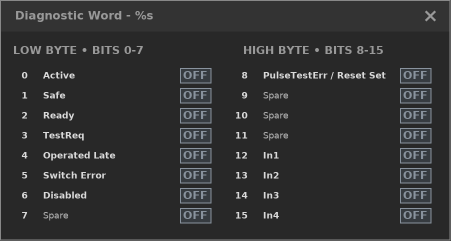
VISUALIZATION FRM_WordDiagnostic  // 451x241
    Rectangle (0,30 451x211)
    Textfield (0,0 411x31), "Diagnostic Word - %s", text variable: Motion_Safety.stSafety.stOut.astDiagnosticElement[GVL_Safety.nHMIDiagWordIndex].sName
    Label (10,40 113x21), "LOW BYTE • BITS 0-7"
    Label (240,40 113x21), "HIGH BYTE • BITS 8-15"
    Label (10,70 21x11), "0"
    Label (10,90 21x11), "1"
    Label (10,110 21x11), "2"
    Label (10,130 21x11), "3"
    Label (10,150 21x11), "4"
    Label (10,170 21x11), "5"
    Label (10,190 21x11), "6"
    Label (10,210 21x11), "7"
    Label (40,70 131x11), "Active"
    Label (40,90 131x11), "Safe"
    Label (40,110 131x11), "Ready"
    Label (40,130 131x11), "TestReq"
    Label (40,150 131x11), "Operated Late"
    Label (40,170 131x11), "Switch Error"
    Label (40,190 131x11), "Disabled"
    Label (40,210 131x11), "Spare"
    Rectangle (180,68 31x15), "ON"
    Rectangle (180,68 31x15), "OFF", invisible if: Motion_Safety.fbMotionSafety.stPNOZEtherCATDiagIn.astDiagnosticElementsIn[GVL_Safety.nHMIDiagWordIndex].nLow.b0
    Rectangle (180,88 31x15), "ON"
    Rectangle (180,88 31x15), "OFF", invisible if: Motion_Safety.fbMotionSafety.stPNOZEtherCATDiagIn.astDiagnosticElementsIn[GVL_Safety.nHMIDiagWordIndex].nLow.b1
    Rectangle (180,108 31x15), "ON"
    Rectangle (180,108 31x15), "OFF", invisible if: Motion_Safety.fbMotionSafety.stPNOZEtherCATDiagIn.astDiagnosticElementsIn[GVL_Safety.nHMIDiagWordIndex].nLow.b2
    Rectangle (180,128 31x15), "ON"
    Rectangle (180,128 31x15), "OFF", invisible if: Motion_Safety.fbMotionSafety.stPNOZEtherCATDiagIn.astDiagnosticElementsIn[GVL_Safety.nHMIDiagWordIndex].nLow.b3
    Rectangle (180,148 31x15), "ON"
    Rectangle (180,148 31x15), "OFF", invisible if: Motion_Safety.fbMotionSafety.stPNOZEtherCATDiagIn.astDiagnosticElementsIn[GVL_Safety.nHMIDiagWordIndex].nLow.b4
    Rectangle (180,168 31x15), "ON"
    Rectangle (180,168 31x15), "OFF", invisible if: Motion_Safety.fbMotionSafety.stPNOZEtherCATDiagIn.astDiagnosticElementsIn[GVL_Safety.nHMIDiagWordIndex].nLow.b5
    Rectangle (180,188 31x15), "ON"
    Rectangle (180,188 31x15), "OFF", invisible if: Motion_Safety.fbMotionSafety.stPNOZEtherCATDiagIn.astDiagnosticElementsIn[GVL_Safety.nHMIDiagWordIndex].nLow.b6
    Rectangle (180,208 31x15), "ON"
    Rectangle (180,208 31x15), "OFF", invisible if: Motion_Safety.fbMotionSafety.stPNOZEtherCATDiagIn.astDiagnosticElementsIn[GVL_Safety.nHMIDiagWordIndex].nLow.b7
    Label (230,70 21x11), "8"
    Label (230,90 21x11), "9"
    Label (230,110 21x11), "10"
    Label (230,130 21x11), "11"
    Label (230,150 21x11), "12"
    Label (230,170 21x11), "13"
    Label (230,190 21x11), "14"
    Label (230,210 21x11), "15"
    Label (260,70 131x11), "PulseTestErr / Reset Set"
    Label (260,90 131x11), "Spare"
    Label (260,110 131x11), "Spare"
    Label (260,130 131x11), "Spare"
    Label (260,150 131x11), "In1"
    Label (260,170 131x11), "In2"
    Label (260,190 131x11), "In3"
    Label (260,210 131x11), "In4"
    Rectangle (400,68 31x15), "ON"
    Rectangle (400,68 31x15), "OFF", invisible if: Motion_Safety.fbMotionSafety.stPNOZEtherCATDiagIn.astDiagnosticElementsIn[GVL_Safety.nHMIDiagWordIndex].nHigh.b0
    Rectangle (400,88 31x15), "ON"
    Rectangle (400,88 31x15), "OFF", invisible if: Motion_Safety.fbMotionSafety.stPNOZEtherCATDiagIn.astDiagnosticElementsIn[GVL_Safety.nHMIDiagWordIndex].nHigh.b1
    Rectangle (400,108 31x15), "ON"
    Rectangle (400,108 31x15), "OFF", invisible if: Motion_Safety.fbMotionSafety.stPNOZEtherCATDiagIn.astDiagnosticElementsIn[GVL_Safety.nHMIDiagWordIndex].nHigh.b2
    Rectangle (400,128 31x15), "ON"
    Rectangle (400,128 31x15), "OFF", invisible if: Motion_Safety.fbMotionSafety.stPNOZEtherCATDiagIn.astDiagnosticElementsIn[GVL_Safety.nHMIDiagWordIndex].nHigh.b3
    Rectangle (400,148 31x15), "ON"
    Rectangle (400,148 31x15), "OFF", invisible if: Motion_Safety.fbMotionSafety.stPNOZEtherCATDiagIn.astDiagnosticElementsIn[GVL_Safety.nHMIDiagWordIndex].nHigh.b4
    Rectangle (400,168 31x15), "ON"
    Rectangle (400,168 31x15), "OFF", invisible if: Motion_Safety.fbMotionSafety.stPNOZEtherCATDiagIn.astDiagnosticElementsIn[GVL_Safety.nHMIDiagWordIndex].nHigh.b5
    Rectangle (400,188 31x15), "ON"
    Rectangle (400,188 31x15), "OFF", invisible if: Motion_Safety.fbMotionSafety.stPNOZEtherCATDiagIn.astDiagnosticElementsIn[GVL_Safety.nHMIDiagWordIndex].nHigh.b6
    Rectangle (400,208 31x15), "ON"
    Rectangle (400,208 31x15), "OFF", invisible if: Motion_Safety.fbMotionSafety.stPNOZEtherCATDiagIn.astDiagnosticElementsIn[GVL_Safety.nHMIDiagWordIndex].nHigh.b7
    Rectangle (410,0 41x31), "×"
        OnMouseUp: CloseDialog Dialog=FRM_WordDiagnostic, Result=None, NumpadKeypadSet=True
END_VISUALIZATION

(* stored: Version 1.1.0.1
   Visu FRM_WordDiagnostic: Id {fc01c149-5aa2-0c0d-10c4-876f67fd2aeb} *)
